{attribute 'no_assign'}
FUNCTION_BLOCK FB_DO_WTURBINE_LD0_WROT1_Beh EXTENDS FB_AcsiCommonDataClass
VAR_INPUT
	stVal: FB_AcsiDATypeBeh := (Fc:=ACSI_FC_ST, TrgOp:=ACSI_TrgOp_dchg OR ACSI_TrgOp_dupd, bLinkResult:=THIS^.AddDataToContainer(ipData:=stVal));
	q: FB_AcsiDATypeQuality := (Fc:=ACSI_FC_ST, TrgOp:=ACSI_TrgOp_qchg, bLinkResult:=THIS^.AddDataToContainer(ipData:=q));
	t: FB_AcsiDATypeTimeStamp := (Fc:=ACSI_FC_ST, bLinkResult:=THIS^.AddDataToContainer(ipData:=t));
END_VAR
VAR
END_VAR

END_FUNCTION_BLOCK

(* stored: Version 1.1.0.1
   POU FB_DO_WTURBINE_LD0_WROT1_Beh: Id {7285ce1e-3c10-4391-9d7a-abdbb57eaed3}, SpecialFunc None *)
